(* IEC 61131-3 sources: plc-vscode/tests/st/test-ready/trust-platform/examples/OSCAT/maintenance_stack/non-oop/src, 3 files *)

(* ---- Configuration.st ---- *)
CONFIGURATION MaintenanceStackClassicConfiguration
RESOURCE Cpu0 ON PLC
    TASK MainTask (INTERVAL := T#100ms, PRIORITY := 1);
    PROGRAM Main WITH MainTask : Main;
END_RESOURCE
END_CONFIGURATION

(* ---- Main.st ---- *)
PROGRAM Main
VAR
    WorkStack : STACK_16;
    CurrentWorkOrder : DWORD;
END_VAR

WorkStack(DIN := DWORD#16#2001, E := TRUE, RD := FALSE, WD := TRUE, RST := FALSE);
WorkStack(DIN := DWORD#16#2002, E := TRUE, RD := FALSE, WD := TRUE, RST := FALSE);
WorkStack(DIN := DWORD#0, E := TRUE, RD := TRUE, WD := FALSE, RST := FALSE);
CurrentWorkOrder := WorkStack.DOUT;
END_PROGRAM

(* ---- Tests.st ---- *)
TEST_PROGRAM MaintenanceStackClassicReturnsNewestWorkOrderFirst
VAR
    WorkStack : STACK_16;
END_VAR

WorkStack(DIN := DWORD#0, E := TRUE, RD := FALSE, WD := FALSE, RST := TRUE);
WorkStack(DIN := DWORD#16#2001, E := TRUE, RD := FALSE, WD := TRUE, RST := FALSE);
WorkStack(DIN := DWORD#16#2002, E := TRUE, RD := FALSE, WD := TRUE, RST := FALSE);
WorkStack(DIN := DWORD#0, E := TRUE, RD := TRUE, WD := FALSE, RST := FALSE);

ASSERT_EQUAL(EXPECTED := DWORD#16#2002, ACTUAL := WorkStack.DOUT);
END_TEST_PROGRAM
